// TIA Portal V19 export
DATA_BLOCK "HMI"   // DB5
{ S7_Optimized_Access := 'TRUE' }
// stored: MemoryReserve 100
   VAR
      ManualMode_Bypass : Bool;
      AutoMode_Bypass : Bool;
   END_VAR
BEGIN
END_DATA_BLOCK
